// Diagnostics API/UDS/API/bds_uds_registerDidWriteCallback
///This function registers the callback for DID write operation.
///
///=======
/// Remarks:
///=======
///    + This is the mandatory API to be used if the DID parameter needs to be written.
///    + The |GVL_uds| is given for usage of defines.
///
///----------
/// FFI:
///----------
///This API can be used in trusted partitions only. See Freedom from Interference (FFI) concept for more details.
///
///==================================================================		  			===================================================================================================
///Return value    								  									Description
///==================================================================		  			===================================================================================================
///0																					No error
///1																					Invalid pointer
///
///==================================================================		   			===================================================================================================
///
///=======
///Code Example:
///=======
///============================================================================
///
///FUNCTION POU_1 : BYTE
///VAR_INPUT
///
///    can_data : POINTER TO BYTE;
///END_VAR
///
///VAR
///    data_au8 : ARRAY[0..8] OF BYTE;
///	
///    i1: BYTE;
///	
///    DidValue_u16: UINT;
///	
///    set_u8: USINT;
///END_VAR
///
///
///bds_uds_GetActiveDid(ADR(DidValue_u16));
///
///IF (DidValue_u16=16#100)
///
///  THEN bds_uds_setCallbackStatus(0);(*positive response for DID 16#100*)
///  
///END_IF
///
///IF (DidValue_u16=16#200) 
///
///  THEN  bds_uds_setCallbackStatus(1);(*negative response for DID 16#200*)
///  
///END_IF
///
///
///FOR i1 := 0 TO 8 BY 1 DO
///can_data[i1]  := data_au8[i1];
///END_FOR;
///POU_1 :=1;
///
///(*Registering callback*)
///
///PROGRAM POU_10
///VAR
///
///	flag_1 : BOOL := 1;
///	
///    flag_2 : BOOL := 1; 
///   
///    flag_3 : BOOL := 1;    
///
///END_VAR
///
///IF ( flag_1)
///
///    THEN bds_uds_registerDidReadCallback (ADR(POU_1));
///
///    flag_1 := 0;(*To make api call once in application*)
///
///END_IF
///
///IF ( flag_2)
///
///    THEN bds_uds_registerDidWriteCallback (ADR(POU_1));
///
///    flag_2 := 0;(*To make api call once in application*)
///
///END_IF
///
///IF ( flag_3)
///
///    THEN bds_uds_registerRoutineF000Callback (ADR(POU_3));
///
///    flag_3 := 0;(*To make api call once in application*)
///
///END_IF
///
///
///============================================================================
{attribute 'external_name' := 'cmp_rts_bds_uds_registerDidWriteCallback'}
FUNCTION bds_uds_registerDidWriteCallback : USINT
VAR_INPUT
	///Function pointer with argument of UINT8 data pointer
	func_pf: POINTER TO BOOL;
END_VAR

END_FUNCTION

// Diagnostics API/UDS/API/bds_uds_registerRoutineF000Callback
///This function will registers the callback for the routine control identifier F000.
///
///=======
/// Remarks:
///=======
///    + This is the mandatory API to be used for routine control identifier F000.
///	+ This is the common register API for routine control F000 for all sub functions like start(), stop(), getResults().
///    + The |GVL_uds| is given for usage of defines.
///
///----------
/// FFI:
///----------
///This API can be used in trusted partitions only. See Freedom from Interference (FFI) concept for more details.
///
///==================================================================		  			===================================================================================================
///Return value    								  									Description
///==================================================================		  			===================================================================================================
///0																					No error
///1																					Invalid pointer
///
///==================================================================		   			===================================================================================================
///
///=======
///Code Example:
///=======
///============================================================================
///
///FUNCTION POU_3 : BYTE
///VAR_INPUT
///
///    dataIn1 : BYTE;
///
///    status : BYTE;
///
///    dataOut1 : POINTER TO BYTE;
///
///    Error_Code : POINTER TO BYTE;
///
///    subservice_u8 : BYTE;
///END_VAR
///
///VAR
///    data_au8: ARRAY[0..7] OF BYTE :=[1,2,3,4,5,6,7,8];
///
///    i: BYTE;
///
///    RidValue_u16: UINT;
///
///    set: BYTE;
///END_VAR
///
///IF(subservice_u8=1)
///
///    THEN bds_uds_setCallbackStatus(0);
///
///END_IF
///
///IF(subservice_u8=2)
///
///    THEN bds_uds_setCallbackStatus(0);
///
///END_IF
///
///IF(subservice_u8=3)
///
///    THEN bds_uds_setCallbackStatus(1);
///
///END_IF
///
///(*Registering callback*)
///
///PROGRAM POU_10
///VAR
///   
///    flag_3 : BOOL := 1;    
///
///END_VAR
///
///
///IF ( flag_3)
///
///    THEN bds_uds_registerRoutineF000Callback (ADR(POU_3));
///
///    flag_3 := 0;(*To make api call once in application*)
///
///END_IF
///
///
///============================================================================
{attribute 'external_name' := 'cmp_rts_bds_uds_registerRoutineF000Callback'}
FUNCTION bds_uds_registerRoutineF000Callback : USINT
VAR_INPUT
	///Function pointer with argument of as mentioned above
	func_pf: POINTER TO BOOL;
END_VAR

END_FUNCTION

// Diagnostics API/UDS/API/bds_uds_getActiveSession
///This function gets the active session of the server/ECU.
///
///=======
/// Remarks:
///=======
///    + By default the server/ECU will be in the Default session after startup.
///    + The |GVL_uds| is given for usage of defines.
///
///----------
/// FFI:
///----------
///This API can be used in trusted partitions. For untrusted partitions use |bds_uds_getActiveSession_ffi|. See Freedom from Interference (FFI) concept for more details.
///
///==================================================================		  			===================================================================================================
///Return value    								  									Description
///==================================================================		  			===================================================================================================
///16#00																				No error
///16#01																				Invalid pointer
///16#25																				FFI API access error.
///
///==================================================================		   			===================================================================================================
///=======
///Code Example:
///=======
///============================================================================
///
///PROGRAM PLC_PRG
///  VAR
///  
///	bds_uds_session_u8:USINT;
///
///	result: USINT;
///	
///  END_VAR
///
///  (*get the active session of the ECU*)
///  
///result := bds_uds_getActiveSession(ADR(bds_uds_session_u8));
///
///============================================================================
{attribute 'external_name' := 'cmp_rts_bds_uds_getActiveSession'}
FUNCTION bds_uds_getActiveSession : USINT
VAR_INPUT
	///Reference of variable where the active session will be saved by the API. 
	///
	///The possible values are:
	///    + DEFAULT SESSION - 16#01
	///    + PROGRAMMING SESSION - 16#02
	///    + EXTENDED DIAGNOSTIC SESSION - 16#03
	///    + SAFETY SYSTEM DIAGNOSTIC SESSION - 16#04
	///    + EOL SESSION - 16#40
	bds_uds_session_u8: POINTER TO USINT;
END_VAR

END_FUNCTION

// Diagnostics API/UDS/FFI_API/bds_uds_getActiveSession_ffi
{attribute 'external_name' := 'cmp_rts_bds_uds_getActiveSession_ffi'}
FUNCTION bds_uds_getActiveSession_ffi : USINT
VAR_INPUT
	///Reference of variable where the active session will be saved by the API. 
	///
	///The possible values are:
	///    + DEFAULT SESSION - 16#01
	///    + PROGRAMMING SESSION - 16#02
	///    + EXTENDED DIAGNOSTIC SESSION - 16#03
	///    + SAFETY SYSTEM DIAGNOSTIC SESSION - 16#04
	///    + EOL SESSION - 16#40
	bds_uds_session_u8: POINTER TO USINT;
END_VAR

END_FUNCTION

// Diagnostics API/UDS/API/bds_uds_getNodeID
///This function reads the currently configured node ID, tester ID and RX/TX identifier from UDS stack and updates the input parameter.
///
///=======
/// Remarks:
///=======
///    + This function reads the UDS parameters of BODAS instance.
///    + The |GVL_uds| is given for usage of defines.
///
///----------
/// FFI:
///----------
///This API can be used in trusted partitions. For untrusted partitions use |bds_uds_getNodeID_ffi|. See Freedom from Interference (FFI) concept for more details.
///		
///==================================================================		  			===================================================================================================
///Return value    								  									Description
///==================================================================		  			===================================================================================================
///16#00																				No error
///16#01																				Node ID read failed
///16#02																				Invalid parameter
///16#25																				FFI API access error.
///
///==================================================================		   			===================================================================================================
{attribute 'external_name' := 'cmp_rts_bds_uds_getNodeID'}
FUNCTION bds_uds_getNodeID : USINT
VAR_INPUT
	///This is a union of a structure and UDINT variable.Default value : 
	///    + nodeid_u8 = 16#01
	///    + testerid_u8 = 16#FA
	///    + rxtxidentifiers_u16 = 16#18DA
	udsConfig_u: POINTER TO bds_uds_udsconfigparameter_tu;
END_VAR

END_FUNCTION

// Diagnostics API/UDS/FFI_API/bds_uds_getNodeID_ffi
{attribute 'external_name' := 'cmp_rts_bds_uds_getNodeID_ffi'}
FUNCTION bds_uds_getNodeID_ffi : USINT
VAR_INPUT
	///This is a union of a structure and UDINT variable.Default value : 
	///    + nodeid_u8 = 16#01
	///    + testerid_u8 = 16#FA
	///    + rxtxidentifiers_u16 = 16#18DA
	udsConfig_u: POINTER TO bds_uds_udsconfigparameter_tu;
END_VAR

END_FUNCTION

// Diagnostics API/UDS/API/bds_uds_permitAccess
///This function sets the access related to the BODAS-service features.
///
///=======
/// Remarks:
///=======
///    + This function needs to be called if access to the BODAS-service to be prevented/permitted.
///    + By default all the services of the BODAS-service is allowed by the BSW.
///    + Multiple bits can be set at a time.
///    + The |GVL_uds| is given for usage of defines.
///
///-----
/// DANGER:
///-----
///
///Application should take care of Programming session bit carefully.
///
///----------
/// FFI:
///----------
///This API can be used in trusted partitions only. See Freedom from Interference (FFI) concept for more details.
///
///==================================================================		  			===================================================================================================
///Return value    								  									Description
///==================================================================		  			===================================================================================================
///0																					No error
///1																					Invalid pointer
///
///==================================================================		   			===================================================================================================
///=======
///Code Example:
///=======
///============================================================================
///
///PROGRAM PLC_PRG
///  VAR
///
///	bds_uds_access_u8:USINT:=0;	
///
///	result: USINT;
///	
///  END_VAR
///  
///result:=bds_uds_permitAccess(bds_uds_access_u8);
///
///============================================================================
{attribute 'external_name' := 'cmp_rts_bds_uds_permitAccess'}
FUNCTION bds_uds_permitAccess : USINT
VAR_INPUT
	///This value defines the coded access rights for the diagnostics services of BODAS-service.
	///	
	///The supported values are:
	///    + 16#00: Prevent all services by BODAS-service.
	///    + 16#01: Permit soft reset by BODAS-service.
	///    + 16#02: Permit hard reset by BODAS-service.
	///    + 16#04: Permit keyOffOn reset by BODAS-service.
	///    + 16#10: Permit to programming session by BODAS-service.
	///    + 16#FF: Permit all services by BODAS-service. (Default)
	bds_uds_access_u8: USINT;
END_VAR

END_FUNCTION

// Diagnostics API/UDS/API/bds_uds_registerRoutineCtrlCallback
///This function will registers the callback for the any routine control configured in easyConfig.
///
///=======
/// Remarks:
///=======
///    + This API is not used for routine control identifier F000. see |bds_uds_registerRoutineF000Callback|
///	+ This is the common register API for all routine control for all sub functions like start(), stop(), getResults().
///    + The |GVL_uds| is given for usage of defines.
///
///----------
/// FFI:
///----------
///This API can be used in trusted partitions only. See Freedom from Interference (FFI) concept for more details.
///
///==================================================================		  			===================================================================================================
///Return value    								  									Description
///==================================================================		  			===================================================================================================
///0																					No error
///1																					Invalid pointer
///
///==================================================================		   			===================================================================================================
///
///=======
///Code Example:
///=======
///============================================================================
///
///FUNCTION POU_3 : BYTE
///VAR_INPUT
///
///    dataIn1 : POINTER TO BYTE;
///
///    status : BYTE;
///
///    dataOut1 : POINTER TO BYTE;
///
///    Error_Code : POINTER TO BYTE;
///
///	(*subservice not available for this function*)
///
///END_VAR
///
///VAR
///    data_au8: ARRAY[0..7] OF BYTE :=[1,2,3,4,5,6,7,8];
///
///    i: BYTE;
///
///    RidValue_u16: UINT;
///
///    set: BYTE;
///END_VAR
///
///IF(subservice_u8=1) THEN
///
///     bds_uds_setCallbackStatus(0);
///
///END_IF
///
///IF(subservice_u8=2) THEN
///
///     bds_uds_setCallbackStatus(0);
///
///END_IF
///
///IF(subservice_u8=3) THEN
///
///     bds_uds_setCallbackStatus(1);
///
///END_IF
///
///(*Registering callback*)
///
///PROGRAM POU_10
///VAR
///   
///    flag_3 : BOOL := 1;    
///
///END_VAR
///
///
///IF ( flag_3)
///
///    THEN bds_uds_registerRoutineCtrlCallback (ADR(POU_3));
///
///    flag_3 := 0;(*To make api call once in application*)
///
///END_IF
///
///
///============================================================================
{attribute 'external_name' := 'cmp_rts_bds_uds_registerRoutineCtrlCallback'}
FUNCTION bds_uds_registerRoutineCtrlCallback : USINT
VAR_INPUT
	///Function pointer with argument as mentioned above
	func_pf: POINTER TO BOOL;
END_VAR

END_FUNCTION

// I/O API/OUT_LEGACY/bds_out_po_disableTstPls
///Disables test pulses for a dedicated proportional output to avoid having test pulses for error detection on that output.
///
///=======
/// Remarks:
///=======
///
///   + Test pulses are enabled by default.
///   + For some application the test pulses may disturb the required functionality of an output. For example if you want to use it for power supply.
///   + The test pulses can be deactivated for High Power Outputs only.
///   + This function should be called only once in the application.
///
///----------
/// FFI:
///----------
///This API can be used in trusted partitions . For untrusted partitions use |bds_out_po_disableTstPls_ffi|. See Freedom from Interference (FFI) concept for more details.
///
///------
/// Attention:
///------
///
///If test pulses are disabled for an output, fault detection and healing is limited.
///
///==================================================================		  			===================================================================================================
///Return value    								  									Description
///==================================================================		  			===================================================================================================
///0																					No error.
///1																					Signal is out of range.
///2																					State Command out of range.
///3																					Output is configured as safout, Test pulse can't be disabled
///
///==================================================================		   			===================================================================================================
///
///=======
///Code Example:
///=======
///============================================================================
///
///PROGRAM PLC_PRG
///
///VAR
///
///	Init_flag_u8:USINT:=0;
///
///END_VAR
///  
///IF(Init_flag_u8=0) THEN (*To make api call once in application*)
///				
///	(* disable test pulses for output K07 *)
///	
///	bds_out_po_disableTstPls(bds_out_po_signal_te.K07, STD_ON);
///  
///	Init_flag_u8:=1;
///  
///END_IF
///
///============================================================================
{attribute 'external_name' := 'cmp_rts_bds_out_po_disableTstPls'}
FUNCTION bds_out_po_disableTstPls : USINT
VAR_INPUT
	///The connector assigned signal name of the output.
	signal_e: UINT;
	///The states are
	///   + STD_OFF - Enables the test pulses (default)
	///   + STD_ON   - Disables the test pulses
	state_u8: USINT;
END_VAR

END_FUNCTION

// I/O API/OUT/FFI_API/bds_out_po_disableTstPls_ffi
{attribute 'external_name' := 'cmp_rts_bds_out_po_disableTstPls_ffi'}
FUNCTION bds_out_po_disableTstPls_ffi : USINT
VAR_INPUT
	///The connector assigned signal name of the output.
	signal_e: UINT;
	///The states are
	///   + STD_OFF - Enables the test pulses (default)
	///   + STD_ON   - Disables the test pulses
	state_u8: USINT;
END_VAR

END_FUNCTION

// I/O API/OUT_LEGACY/bds_out_po_getCurrent
///Get the current of the proportional output.
///
///=======
/// Remarks:
///=======
///   + The threshold for the over current detection is 6000mA and therefore also the measurement range is defined from 0..6000mA.
///
///----------
/// FFI:
///----------
///This API can be used in trusted partitions . For untrusted partitions use |bds_out_po_getCurrent_ffi|. See Freedom from Interference (FFI) concept for more details.
///
///==================================================================		  			===================================================================================================
///Return value    								  									Description
///==================================================================		  			===================================================================================================
///0																					No error.
///1																					A parameter is invalid.
///2																					Function call was erroneous.
///
///==================================================================		   			===================================================================================================
///
///=======
///Code Example:
///=======
///============================================================================
///
///PROGRAM appl_10ms_task
///VAR
///bds_outClcU_signal_e : bds_outClcU_signal_te;
/// bds_outClcU_retSetVoltage_s : bds_outClcU_setVoltage_ts;
/// u_mV_u16 : UINT := 8000;
///END_VAR
///
///bds_outClcU_signal_e := bds_outClcU_K62_E;
///
///bds_outClcU_retSetVoltage_s := bds_outClcU_setVoltage(bds_outClcU_signal_e, u_mV_u16);
///
///IF bds_outCmn_ok_E = bds_outClcU_retSetVoltage_s.statusApi_e THEN
/// (* Call successful, signal is valid )
/// ( Set point value is set on requested output )
///  ELSE
///  ( error handling *)
///  END_IF
///
///END_PROGRAM
///============================================================================
{attribute 'external_name' := 'cmp_rts_bds_out_po_getCurrent'}
FUNCTION bds_out_po_getCurrent : USINT
VAR_INPUT
	///The connector assigned signal name of the output.
	signal_e: UINT;
	///Storage address of the value.
	///
	///   + Range:0 to 60000 [mA]
	value_pu16: POINTER TO UINT;
END_VAR

END_FUNCTION

// I/O API/OUT/FFI_API/bds_out_po_getCurrent_ffi
{attribute 'external_name' := 'cmp_rts_bds_out_po_getCurrent_ffi'}
FUNCTION bds_out_po_getCurrent_ffi : USINT
VAR_INPUT
	///The connector assigned signal name of the output.
	signal_e: UINT;
	///Storage address of the value.
	///
	///   + Range:0 to 60000 [mA]
	value_pu16: POINTER TO UINT;
END_VAR

END_FUNCTION

// I/O API/OUT/API/bds_outClcU_setVoltage
///The BODAS API-Function sets the analog voltage set point of the output signal.
///
///=======
/// Remarks:
///=======
///    +For AOV analog voltage output the set voltage range is from 0 to 10000mV  (available signal refer to table "AOV Analog Voltage Output" in RC27-18/40 - Outputs).
///    
///    +For PVG proportional voltage output the accepted set voltage range is from 0 to 27000mV (75% of max Ubat) (available signal refer to table "PVG Proportional Voltage Output" in RC27-18/40 - Outputs).
///   
///    +·If the set point has been set to 0 value then the output can also be used as analog voltage input, refer to bds_outClcU_get.
///
///----------
/// FFI:
///----------
///This API can be used in trusted partitions. For untrusted partitions use bds_outClcU_setVoltage_ffi. See Freedom from Interference (FFI) concept for more details.
///
///------
/// Info:
///------
///
/// +For the output type PVG: 
///   
///   +An external load is mandatory, refer to Technical Data Sheet (RE-sheet RE95207).
///   
///   +If the requested voltage set point is higher than 75% of the max possible battery voltage (36V) the return value of the status API function call is: bds_outCmn_outOfRng_E.
///   
///   +·The possible voltage range that can be controlled is 25% to 75% of the actual battery voltage, because of hardware limitations. The internal set point of the regulation will be dynamically limited to this min or max value without setting any error or status information.
///
///   +Example 1: 
///   +Actual battery voltage = 24V and output voltage is set to 4V => results in output voltage = 6V (25% of actual battery voltage).
///
///   +Example 2: 
///   +Actual battery voltage = 12V and output voltage is set to 4V => results in output voltage = 4V (33% of actual battery voltage).
///   
///   +The set point request of 0V is also valid and will switch off the output. 
///   
///   
///   +Macro define "bds_outClcU_strtNumSigAov_D" in easyConfig generated file "bds_outClcU_ec.h" defines the start of the Analog voltage output (AOV) signals in the enumeration type definition "bds_outClcU_signal_te".
///
///
///==================================================================		  			===================================================================================================
///Return value    								  									Description
///==================================================================		  			===================================================================================================
///bds_outClcU_setVoltage_ts															 The return structure containing the state information (statusApi_e)
///
///==================================================================		   			===================================================================================================
///
///=======
///Code Example:
///=======
///============================================================================
///
///PROGRAM appl_10ms_task
///
///VAR
///
///bds_outClcU_signal_e : bds_outClcU_signal_te;
///
///bds_outClcU_retSetVoltage_s : bds_outClcU_setVoltage_ts;
///
///u_mV_u16 : UINT := 8000;
///
///END_VAR
///
///bds_outClcU_signal_e := bds_outClcU_signal_te.bds_outClcU_K62_E;
///
///bds_outClcU_retSetVoltage_s := bds_outClcU_setVoltage(bds_outClcU_signal_e, u_mV_u16);
///
///IF bds_outCmn_ok_E = bds_outClcU_retSetVoltage_s.statusApi_e THEN
///
///(* Call successful, signal is valid *)
///(* Set point value is set on requested output *)
///
///ELSE
///
///(* error handling *)
///
///END_IF
///
///END_PROGRAM
///
///============================================================================
{attribute 'external_name' := 'cmp_rts_bds_outClcU_setVoltage'}
FUNCTION bds_outClcU_setVoltage : bds_outClcU_setVoltage_ts
VAR_INPUT
	///signal name of the output (connector pin)
	signal_e: USINT;
	///New set point for PWM [0.1%] respective AOV [mV].Range:
	///   + PWM: 0 and 250 to 750
	///   + AOV: 0 to 10000
	u_mV_u16: UINT;
END_VAR

END_FUNCTION

// I/O API/OUT/API/bds_outClcU_get
///The BODAS API-Function gets the measured voltage in [mV] of the analog voltage output pin.
///
///=======
/// Remarks:
///=======
///  +The voltage range depends on the type.
/// 
///     +AOV: 0 to 12000mV
/// 
///     +PVG: 0 to 33000mV.
/// 
///  +The read-back path of the analoge voltage can also be used as analog input, if the set point is set to zero, refer also bds_outClcU_setVolatge and bds_outClcU_setPercUBat.
///  +Diagnostics capabilities similar to standard inputs is not available. 
/// 
///  +The status data holds all relevant information of the analog voltage output, see example below.
/// 
///  +Part of the status bit field is also the fault error status of every DFC (e.g. stErrSCB_b1), see topic Digital outputs and Diagnostic Fault Check. 

///
///----------
/// FFI:
///----------
///This API can be used in both trusted and untrusted partitions. See Freedom from Interference (FFI) concept for more details.
///
///------
/// Info:
///------
///
///   +For the predefined pin type analog voltage output (AOV) there is an option in easyConfig tool to reconfigure it as analog voltage input or digital input
///
///
///==================================================================		  			===================================================================================================
///Return value    								  									    Description
///==================================================================		  			===================================================================================================
///bds_outClcU_get_ts															        The return structure containing the measured voltage in [mV] and the state information (statusApi_e)
///
///==================================================================		   			===================================================================================================
///
///=======
///Code Example:
///=======
///============================================================================
///
/// PROGRAM appl_10ms_task 
///
/// VAR
/// 
/// bds_outClcU_signal_e : bds_outClcU_signal_te; 
/// 
/// bds_outClcU_retGet_s : bds_outClcU_get_ts; 
///
/// retVal_uAct_mV_u16, retVal_uSet_mV_u16 : UINT;
/// 
/// END_VAR
///
/// bds_outClcU_signal_e := bds_outClcU_signal_te.bds_outClcU_K62_E; 
///
///
/// (* call BDS-Function - Set voltage output *)
///
/// bds_outClcU_setVoltage(bds_outClcU_signal_e, 8000); 
///
/// (* call BDS-Function - Get status and diagnostic information *)
///
/// bds_outClcU_retGet_s := bds_outClcU_get(bds_outClcU_signal_e); 
///
///
/// IF bds_outCmn_ok_E = bds_outClcU_retGet_s.statusApi_e THEN
///
/// (* Call successful, signal is valid *)
///
/// 	(* check if there is a short cut to battery or to ground? *)
///
///		IF (TRUE = bds_outClcU_retGet_s.statusDiag_b.stErrSCB_b1) OR (TRUE = bds_outClcU_retGet_s.statusDiag_b.stErrSCG_b1) THEN
///
/// 	(* SCB or SCG - Set values to zero *)
///
///  	retVal_uAct_mV_u16 := 0; 
///
/// 	retVal_uSet_mV_u16 := 0; 
///
/// 	ELSE (* get actual measured voltage on requested output *)
///
///		retVal_uAct_mV_u16 := bds_outClcU_retGet_s.uAct_mV_u16; 
///
///     (* get requested set point voltage on requested output *)
///
///     retVal_uSet_mV_u16 := bds_outClcU_retGet_s.uSet_mV_u16; 
///
/// 	END_IF
///
/// ELSE
///
/// (* error handling *)
///
/// END_IF
///
/// END_PROGRAM
///
///============================================================================
{attribute 'external_name' := 'cmp_rts_bds_outClcU_get'}
FUNCTION bds_outClcU_get : bds_outClcU_get_ts
VAR_INPUT
	///signal name of the output (connector pin)
	signal_e: USINT;
END_VAR

END_FUNCTION

// I/O API/OUT/API/bds_outClcU_setPercUBat
/// The BODAS API-Function sets the analog voltage output in percentage value of the the battery voltage.
///
///=======
/// Remarks:
///=======
///    +Set the voltage range FROM 0 AND 250…750 [0.1%] OF the battery voltage OF the PVG analog voltage output (available signal refer TO table "PVG Proportional Voltage Output" in RC27-18/40 - Outputs).

///    +If the set point has been set to 0 value then the output can also be used as analog voltage input, refer to bds_outClcU_get.

///
///----------
/// FFI:
///----------
/// This API can be used in trusted partitions. For untrusted partitions use bds_outClcU_setPercUBat_ffi. See Freedom from Interference (FFI) concept for more details.
///
///------
/// Info:
///------
///
/// +For the output type PVG an external load is mandatory, refer to Technical Data Sheet (RE-sheet RE95207).
/// +Macro define "bds_outClcU_strtNumSigAov_D" in easyConfig generated file "bds_outClcU_ec.h" defines the start of the Analog voltage output (AOV) signals in the enumeration type definition "bds_outClcU_signal_te"
///
///
///==================================================================		  			===================================================================================================
///Return value    								  									    Description
///==================================================================		  			===================================================================================================
///bds_outClcU_setPercUBat_ts														     The return structure containing the state information (statusApi_e)
///
///==================================================================		   			===================================================================================================
///
///=======
///Code Example:
///=======
///============================================================================
///
/// PROGRAM appl_10ms_task 
///
/// VAR bds_outClcU_signal_e : bds_outClcU_signal_te;
///
/// bds_outClcU_retSetPercUBat_s : bds_outClcU_setPercUBat_ts;
///
/// ratUBat_perml_u16 : UINT;
///
/// END_VAR
///
/// bds_outClcU_signal_e := bds_outClcU_signal_te.bds_outClcU_K25_E;
///
/// ratUBat_perml_u16 := 750;
///
///bds_outClcU_retSetPercUBat_s := bds_outClcU_setPercUBat(bds_outClcU_signal_e, ratUBat_perml_u16);
///
///IF bds_outCmn_ok_E = bds_outClcU_retSetPercUBat_s.statusApi_e THEN 
///
/// (* Call successful, signal is valid *)
///
/// (* Set point value is set on requested output *)
///
/// ELSE
/// 
/// (* error handling *)
///
/// END_IF
///
/// END_PROGRAM
///
///============================================================================
{attribute 'external_name' := 'cmp_rts_bds_outClcU_setPercUBat'}
FUNCTION bds_outClcU_setPercUBat : bds_outClcU_setPercUBat_ts
VAR_INPUT
	///signal name of the output (connector pin)
	signal_e: USINT;
	///voltage set point in 0, 250...750 [0.1%] of battery voltage
 
	ratUBat_perml_u16: UINT;
END_VAR

END_FUNCTION

// Diagnostics API/UDS/API/bds_uds_setUUID
///This function is to set the Universal Unique Identifier for ODX file data identification.
///
///=======
/// Remarks:
///=======
///
///    + UDS dataidentifier 16#F19E supports the UUID-ODX data identification value set from |bds_uds_setUUID|.
///    + The |GVL_uds| is given for usage of defines.
///    + This API should be called once in Application
///
///----------
/// FFI:
///----------
///This API can be used in trusted partitions only. See Freedom from Interference (FFI) concept for more details.
///
///----------
/// WARNING:
///----------
///
///This function should be called only once in the application.
///
///==================================================================		  			===================================================================================================
///Return value    								  									Description
///==================================================================		  			===================================================================================================
///16#00																				No error
///16#01																				Invalid pointer
///
///==================================================================		   			===================================================================================================
///=======
///Code Example:
///=======
///============================================================================
///
///PROGRAM PLC_PRG
///  VAR
///
///	bds_uds_uuid_pu8: ARRAY[0 .. 17] OF USINT;
///
///	bds_uds_uuidLen_u8 : USINT := 18;
///
///	result: USINT;
///
///	FLAG: BOOL;
///	
///  END_VAR
///  
///IF FLAG:=FALSE THEN
///
///	bds_uds_uuid_pu8[0]:= 16#FF; 
///
///	bds_uds_uuid_pu8[1]:= 16#AA; 
///
///	result := bds_uds_setUUID(ADR(bds_uds_uuid_pu8),bds_uds_uuidLen_u8);
///
///	FLAG:= TRUE;
///
///END_IF
///
///============================================================================
{attribute 'external_name' := 'cmp_rts_bds_uds_setUUID'}
FUNCTION bds_uds_setUUID : USINT
VAR_INPUT
	///Array index for the 18 byte UUID value for ODX identification
	bds_uds_uuid_pu8: POINTER TO USINT;
	///Length in bytes for the UUID value, maximum is 18.
	bds_uds_uuidLen_u8: USINT;
END_VAR

END_FUNCTION

// I/O API/SAFOUT/API/bds_safout_cfgDiag
///Configures the allowed current deviation limit for current deviation monitoring between high side and low side outputs of a safout channel. 
///
///=======
/// Remarks:
///=======
///   + The allowed default current deviation limit is 100 mA. Current deviation monitoring between high side and low side outputs is supported only for PHMDL, PLMDH, PLDHS and PHDLS mode.
///   + Some of the errors are detected using current deviation monitoring, setting of allowed current deviation limit shall be chosen wisely for the application. 
///   + Total allowed current deviation limit = (Current deviation in mA + (percentage of sum of current through multiple side outputs in previous100 ms) in mA).
///
///----------
/// FFI:
///----------
///This API can be used in trusted partitions only. See Freedom from Interference (FFI) concept for more details.
///
///------
/// CAUTION:
///------
///
///Be careful while configuring current deviation.
///
///==================================================================		  			===================================================================================================
///Return value    								  									Description
///==================================================================		  			===================================================================================================
///0																					No error
///1																					A parameter is invalid
///2																					Wrong mode or channel
///3																					Feature not supported for safout mode
///
///==================================================================		   			===================================================================================================
///
///=======
///Code Example:
///=======
///============================================================================
///
///VAR_GLOBAL CONSTANT
///
///   (* safout channel name *)
///
///   PHDLS_CHNL1: UINT := (PHDLS OR CHNL1);
///
///   DHDLM_CHNL2: UINT := (DHDLM OR CHNL2);
///
///   PHMDL_CHNL3: UINT := (PHMDL OR CHNL3);
///   
///   PLDHS_CHNL4: UINT := (PLDHS OR CHNL4);
///
///   DLDHM_CHNL5: UINT := (DLDHM OR CHNL5);
///
///   PLMDH_CHNL6: UINT := (PLMDH OR CHNL6);
///
///END_VAR
///
///PROGRAM PLC_PRG
///
///VAR
///
///END_VAR
///
///
///(* configure for POC *)
///
///bds_out_po_cfg(bds_out_po_signal_te.K73, STD_ACTIVE);
///
///bds_out_po_cfg(bds_out_po_signal_te.K07, STD_ACTIVE);
///
///bds_out_po_cfg(bds_out_po_signal_te.K29, STD_ACTIVE);
///
///bds_out_po_cfg(bds_out_po_signal_te.K09, STD_ACTIVE);
///
///
///
///(* configure channels for SAFOUT *)
///
///bds_safout_cfg(PHDLS_CHNL1, bds_out_po_signal_te.K73, bds_out_po_signal_te.K51, bds_out_do_signal_te.K14, 0, 0);
///
///bds_safout_cfg(DHDLM_CHNL2, bds_out_po_signal_te.K08, bds_out_do_signal_te.K16, bds_out_do_signal_te.K15, bds_out_do_signal_te.K13, 0);
///
///bds_safout_cfg(PHMDL_CHNL3, bds_out_do_signal_te.K12, bds_out_po_signal_te.K07, bds_out_po_signal_te.K29, bds_out_po_signal_te.K09, 0);
///
///bds_safout_cfg(PLDHS_CHNL4, bds_out_po_signal_te.A19, bds_out_po_signal_te.A32, bds_out_do_signal_te.A47, 0, 0);
///
///bds_safout_cfg(DLDHM_CHNL5, bds_out_po_signal_te.A03, bds_out_do_signal_te.A33, bds_out_do_signal_te.A46, bds_out_do_signal_te.A48, 0);
///
///bds_safout_cfg(PLMDH_CHNL6, bds_out_do_signal_te.A31, bds_out_po_signal_te.A05, bds_out_po_signal_te.A20, 0, 0);
///
///bds_safout_cfgDiag(PHDLS_CHNL1, 150,0);
///
///bds_safout_cfgDiag(PHMDL_CHNL3, 200, 10);
///
///bds_safout_cfgDiag(PLDHS_CHNL4, 200,15);
///
///bds_safout_cfgDiag(PLMDH_CHNL6, 200, 10);
///
///============================================================================
{attribute 'external_name' := 'cmp_rts_bds_safout_cfgDiag'}
FUNCTION bds_safout_cfgDiag : USINT
VAR_INPUT
	///The connector assigned signal name of the output.
	///
	///The channel name is composed of mode and channel number
	///
	///channel name = mode OR channel number
	///
	///and shall be defined from the application (see also example below):
	///
	///PHDLS_CHNL1: UINT := (PHDLS OR CHNL1)
	chnl_u16: UINT;
	///Fixed allowed current deviation [mA] 
	///   + Range: 100..1000 
	deviation_u16: UINT;
	///Percentage of allowed current deviation [%]
	///   + Range:0..100
	devPercentage_u8: USINT;
END_VAR

END_FUNCTION

// I/O API/SAFOUT/API/bds_safout_enableTest
///Enables test for Safout channel.
///
///When safout channel is inactive i.e all highsides and lowside are OFF, every 2 seconds a test is performed by switching ON common side for 120 ms.  During test, open load error diagnostic is performed on multiple outputs of the safout channel can be detected.
///
///=======
/// Remarks:
///=======
///   + A channel shall be configured with ECU specific modes, see Safety outputs.
///   + By default, test is disabled 
///   + This test is not performed when there a SCB on HS output / SCG on LS outputs.
///   + Test status can be using |bds_safout_getStatus| API. Test complete flag is reset once status is read by |bds_safout_getStatus|.
///   + This only supported for PHMDL mode. In other safout modes open load is detected without this test.
///
///----------
/// FFI:
///----------
///This API can be used in trusted partitions only. See Freedom from Interference (FFI) concept for more details.
///
///==================================================================		  			===================================================================================================
///Return value    								  									Description
///==================================================================		  			===================================================================================================
///0																					No error.
///1																					A parameter is invalid.
///2																					Not supported for this mode
///
///==================================================================		   			===================================================================================================
///
///=======
///Code Example:
///=======
///============================================================================
///
///VAR_GLOBAL CONSTANT
///
///   (* safout channel name *)
///
///   PHDLS_CHNL1: UINT := (PHDLS OR CHNL1);
///
///   DHDLM_CHNL2: UINT := (DHDLM OR CHNL2);
///
///   PHMDL_CHNL3: UINT := (PHMDL OR CHNL3);
///
///END_VAR
///
///PROGRAM PLC_PRG
///
///VAR
///
///END_VAR
///
///(* configure for POC *)
///
///bds_out_po_cfg(bds_out_po_signal_te.K73, STD_ACTIVE);
///
///bds_out_po_cfg(bds_out_po_signal_te.K07, STD_ACTIVE);
///
///bds_out_po_cfg(bds_out_po_signal_te.K29, STD_ACTIVE);
///
///bds_out_po_cfg(bds_out_po_signal_te.K09, STD_ACTIVE);
///
///
///(* configure channels for SAFOUT *)
///
///bds_safout_cfg(PHDLS_CHNL1, bds_out_po_signal_te.K73, bds_out_po_signal_te.K51, bds_out_do_signal_te.K14, 0, 0);
///
///bds_safout_cfg(DHDLM_CHNL2, bds_out_po_signal_te.K08, bds_out_do_signal_te.K16, bds_out_do_signal_te.K15, bds_out_do_signal_te.K13, 0);
///
///bds_safout_cfg(PHMDL_CHNL3, bds_out_do_signal_te.K12, bds_out_po_signal_te.K07, bds_out_po_signal_te.K29, bds_out_po_signal_te.K09, 0);
///
///bds_safout_enableTest(PHMDL_CHNL3,STD_ON);
///
///============================================================================
{attribute 'external_name' := 'cmp_rts_bds_safout_enableTest'}
FUNCTION bds_safout_enableTest : USINT
VAR_INPUT
	///The connector assigned signal name of the output.
	///
	///The channel name is composed of mode and channel number
	///
	///channel name = mode OR channel number
	///
	///and shall be defined from the application (see also example below):
	///
	///PHDLS_CHNL1: UINT := (PHDLS OR CHNL1)
	chnl_u16: UINT;
	///The states are
	///   + STD_OFF - Disable the test (default)
	///   + STD_ON   - Enable the test
	state_u8: USINT;
END_VAR

END_FUNCTION

// I/O API/IN legacy/API/bds_in_ri_cfg
///Configures the diagnosis threshold resistances for an input. 
///
///=======
/// Remarks:
///=======
///   + The information about definitions and structures can be found in BODAS API library and  bds_rts_ec.xml.
///   + The diagnosis of the input is only possible after the configuration of the thresholds.
///   + With a defined measurement range of 20 to 400k ohm the diagnosis range is defined from 30 to 399.99k ohm.
///   + For more information see |bds_in_ri_getStatus|.
///   + This function should be called only once in the application.
///
///
///----------
/// FFI:
///----------
///This API can be used in trusted partitions only. See Freedom from Interference (FFI) concept for more details.
///
///==================================================================		  			===================================================================================================
///Return value    								  									Description
///==================================================================		  			===================================================================================================
///0																					No error
///1																					Invalid parameter
///2																					Function call was erroneous
///
///==================================================================		   			===================================================================================================
///
///
///=======
///Code Example:
///=======
///============================================================================
///
///PROGRAM PLC_PRG
///
///  VAR
///  
///	Init_flag_u8:USINT:=0;
/// 
///  END_VAR
///  
///IF(Init_flag_u8=0) THEN (*To make api call once in application*)
///
///	(* configure diagnosis thresholds of input K60 *)
///	
///	bds_in_ri_cfg(bds_in_ri_signal_te.K60, 2000, 200);
///	
///	Init_flag_u8:=1;
///  
///END_IF
///
///============================================================================
{attribute 'external_name' := 'cmp_rts_bds_in_ri_cfg'}
FUNCTION bds_in_ri_cfg : USINT
VAR_INPUT
	///The signal name that is assigned to the respective pin configured as resistance input
	signal_e: UINT;
	///Upper diagnosis threshold [ohm].
	///
	///Range: 
	///30 to 399990
	///
	///Note:
	///upperThreshold_u32 > lowerThreshold_u32.  
	upperThreshold_u32: UDINT;
	///Lower diagnosis threshold [ohm].
	///
	///Range: 
	///30 to 399990
	///
	///Note:
	///lowerThreshold_u32 < upperThreshold_u32 
	lowerThreshold_u32: UDINT;
END_VAR

END_FUNCTION

// I/O API/IN legacy/API/bds_in_ri_getStatus
///Provides the status of an input.
///
///=======
/// Remarks:
///=======
///   + For information about the signal acquisition see Analog voltage aquisition.
///   + The status data provides all relevant information of the resistance input.  See the example below.
///	   + A member variable  of  the status data structure  provides the fault status of corresponding  DFC (e.g., stDFC_SCB_u16), see topic Diagnostic Fault Check. 
///	   + With the macros (e.g., bds_dsm_DFC_ldf) defined in bds_dsm_api.h  respective bit fields of the fault status can be read.
///
///----------
/// FFI:
///----------
///This API can be used in trusted partitions only. See Freedom from Interference (FFI) concept for more details.
///
///==================================================================		  			===================================================================================================
///Return value    								  									Description
///==================================================================		  			===================================================================================================
///0																					No error
///1																					Invalid parameter
///
///==================================================================		   			===================================================================================================
///
///=======
///Code Example:
///=======
///============================================================================
///
///PROGRAM appl_10ms_task
///  VAR
///  
///    stK60_s: bds_in_ri_ts;
///	
///    ldf_u8: USINT := 16#00;
///	
///  END_VAR
///
///
///(* get the status of input K60 *)
///
///bds_in_ri_getStatus(bds_in_ri_signal_te.K60, ADR(stK60_s));
///
///  (* get last debounced fault *)
///  
///  ldf_u8 = bds_dsm_DFC_ldf(stK60_s.stDFC_SCB_u16);
///END
///
///============================================================================
{attribute 'external_name' := 'cmp_rts_bds_in_ri_getStatus'}
FUNCTION bds_in_ri_getStatus : USINT
VAR_INPUT
	///The signal name that is assigned to the respective pin configured as resistance input
	signal_e: UINT;
	///Storage address of the data
	data_ps: POINTER TO bds_in_ri_ts;
END_VAR

END_FUNCTION

// I/O API/IN legacy/API/bds_in_ri_cfgTemp
///Configures the resistance inputs for temperature measurement. 
///
///=======
/// Remarks:
///=======
///   + The supported BSW sensors are:
///	   + TSF (sensor type is PTC) 
///	   + TSA (sensor type is PTC)
///	   + TFW (sensor type is NTC)
///   + For additional sensors the corresponding look up tables shall be defined, for more information see Define a look up table for temperature sensors.
///
///
///----------
/// FFI:
///----------
///This API can be used in trusted partitions only. See Freedom from Interference (FFI) concept for more details.
///
///
///==================================================================		  			===================================================================================================
///Return value    								  									Description
///==================================================================		  			===================================================================================================
///0																					No error
///1																					Invalid parameter
///
///==================================================================		   			===================================================================================================
///
///
///=======
///Code Example:
///=======
///============================================================================
///
///PROGRAM PLC_PRG
///
///  VAR
///  
///    lookup_TSF_cau16: ARRAY[1..256] OF UINT := [256(0)];
///	
///    lookup_TSA_cau16: ARRAY[1..256] OF UINT := [256(0)];
///	
///    lookup_TFW_cau16: ARRAY[1..256] OF UINT := [256(0)];
///	
///	Init_flag_u8:USINT:=0;
///	
///  END_VAR
///  
///IF(Init_flag_u8=0) THEN (*To make api call once in application*)
///
///	(* configure temperature sensor of input K60 *)
///	
///	bds_in_ri_cfgTemp(bds_in_ri_signal_te.K60, lookup_TSF_cau16, PTC);
///	
///	bds_in_ri_cfgTemp(bds_in_ri_signal_te.K58, lookup_TFW_cau16, NTC);
///	
///	Init_flag_u8:=1;
///  
///END_IF
///
///============================================================================
{attribute 'external_name' := 'cmp_rts_bds_in_ri_cfgTemp'}
FUNCTION bds_in_ri_cfgTemp : USINT
VAR_INPUT
	///The signal name that is assigned to the respective pin configured as resistance input
	signal_e: UINT;
	///Predefined look up tables for the BODAS-BSW are:
	///   + lookup_TSF_cau16 
	///   + lookup_TSA_cau16
	///   + lookup_TFW_cau16
	lookup_pcau16: POINTER TO UINT;
	///Selected sensor type are:
	///   + NTC 
	///   + PTC 
	type_u8: USINT;
END_VAR

END_FUNCTION

// I/O API/IN legacy/API/bds_in_sent_getSDDatabox
///It provides the oldest slow serial data from a particular databox of a particular SENT channel.
///
///=======
/// Remarks:
///=======
///   + The receive databoxes must be registered with |bds_in_sent_registerSDDataboxes| and then the specific receive databox has to be initialized by |bds_in_sent_initSDDatabox|.
///   + The return value  should be checked first before accessing the data/message.
///
/// 
///----------
/// FFI:
///----------
///This API can be used in trusted partitions only. See Freedom from Interference (FFI) concept for more details.
/// 
///==================================================================		  			===================================================================================================
///Return value    								  									Description
///==================================================================		  			===================================================================================================
///0																					No error
///1																					Invalid parameter
///2																					Databox is not initialized
///3																					Receive buffer is empty
///4																					Receive buffer overflow
///
///==================================================================		   			===================================================================================================
///
///=======
///Code Example:
///=======
///============================================================================
///
///VAR_GLOBAL CONSTANT
///
///   SENT_NUM_DATABOXES_D: USINT := 5;
///
///   SENT_DATABOX_BUFLEN_D: UDINT := 10;
///
///END_VAR
///
/// 
///
///PROGRAM PLC_PRG
///
///   VAR
///
///     sent_dataBox_as: ARRAY[1..SENT_NUM_DATABOXES_D] OF bds_in_sent_SDDataBox_ts;
///
///     sent_slowData1_as: ARRAY[1..SENT_DATABOX_BUFLEN_D] OF bds_in_sent_slowData_ts;
///
///     databoxdata_au16: ARRAY[1..SENT_NUMOFDATABOX_D] OF UINT;
///	 
///	Init_flag_u8:USINT:=0;	 
///
///   END_VAR
///  
///IF(Init_flag_u8=0) THEN (*To make api call once in application*)
///
///   (* register slow databox *)
///
///   bds_in_sent_registerSDDataboxes(bds_in_sent_signal_te.K52, ADR(sent_dataBox_as), SENT_NUM_DATABOXES_D);
///
/// 
///
///   (* initialize the databox *)
///
///   bds_in_sent_initSDDatabox(bds_in_sent_signal_te.K52, 1, 2, ADR(sent_slowData1_as), 5);
///	
///	Init_flag_u8:=1;
///  
///END_IF
///
/// 
///
///PROGRAM appl_10ms_task
///
///  uint8 statusSDDatabox_u8;
///
///  statusSDDatabox_u8 := bds_in_sent_getSDDatabox(bds_in_sent_signal_te.K52,1, &databoxdata_au16[0]);
///
/// 
///
///  IF (0 = statusSDDatabox_u8) THEN
///
///    (* valid data box of SLOW data *)
///
///  END_IF
///
///END
///
///
///============================================================================
{attribute 'external_name' := 'cmp_rts_bds_in_sent_getSDDatabox'}
FUNCTION bds_in_sent_getSDDatabox : USINT
VAR_INPUT
	///The signal name that is assigned to the respective pin configured as SENT input
	signal_e: UINT;
	///Number of data box
	numDatabox_u8: USINT;
	///Pointer to data array
	data_pu16: POINTER TO UINT;
END_VAR

END_FUNCTION

// I/O API/IN legacy/API/bds_in_sent_registerSDDataboxes
///The function registers a slow Databox for a particular message of particular SENT channel. Application has to reserve the memory for databox and databox is managed by the BODAS-BSW.
///
///=======
/// Remarks:
///=======
///
///   + Receive databoxes which has to be registered with function described. Each receive databox has to be initialized with function |bds_in_sent_initSDDatabox|.
///   + The use of receive databoxes is optional.
///   + By default no databoxes are registered. 
///   + For each SENT channel seperate receive databoxes must be registered. 
///   + Please register receive databoxes only as much as needed. Each receive databox increases the system load (if a SENT message is received). 
/// 
///
///----------
/// FFI:
///----------
///This API can be used in trusted partitions only. See Freedom from Interference (FFI) concept for more details.
///
///==================================================================		  			===================================================================================================
///Return value    								  									Description
///==================================================================		  			===================================================================================================
///0																					No error
///1																					Invalid parameter
///2																					new buffer overlaps a present buffer
///
///==================================================================		   			===================================================================================================
///
///=======
///Code Example:
///=======
///============================================================================
///
///VAR_GLOBAL_CONSTANT
///
///   SENT_NUM_DATABOXES_D: USINT := 5;
///
///END_VAR
///
/// 
///
///PROGRAM OsIniProc
///
///   VAR
///
///		sent_dataBox_as: ARRAY[1..SENT_NUM_DATABOXES_D] OF bds_in_sent_SDDataBox_ts;
///		
///		Init_flag_u8:USINT:=0;	 
///
///   END_VAR
///  
///IF(Init_flag_u8=0) THEN (*To make api call once in application*)
///
///	(* register slow databox *)
///	
///	bds_in_sent_registerSDDataboxes(bds_in_sent_signal_te.K57, ADR(sent_dataBox_as), SENT_NUM_DATABOXES_D);
///	
///	Init_flag_u8:=1;
///  
///END_IF
///
///============================================================================
{attribute 'external_name' := 'cmp_rts_bds_in_sent_registerSDDataboxes'}
FUNCTION bds_in_sent_registerSDDataboxes : USINT
VAR_INPUT
	///The signal name that is assigned to the respective pin configured as SENT input
	signal_e: UINT;
	///Pointer to the message data of type |bds_in_sent_SDDataBox_ts|
	mem_pas: POINTER TO bds_in_sent_SDDataBox_ts;
	/// number of receive databoxes
	num_u8: USINT;
END_VAR

END_FUNCTION

// I/O API/IN legacy/API/bds_in_sent_initSDDatabox
///It initializes a slow serial databox for a particular message of a SENT channel. 
///
///=======
/// Remarks:
///=======
///   + The use of receive databoxes is optional.
///   + Before using this function the receive databoxes must be registered with |bds_in_sent_registerSDDataboxes|  
///   + Each receive databox has to be initialized before it can be used.
///   + By default no databoxes are registered. 
///   + Duplication of same ID should be avoided. 
///
///----------
/// FFI:
///----------
///This API can be used in trusted partitions only. See Freedom from Interference (FFI) concept for more details.
///  
///==================================================================		  			===================================================================================================
///Return value    								  									Description
///==================================================================		  			===================================================================================================
///0																					No error
///1																					Invalid parameter
///2																					New buffer overlaps a present buffer
///3																					A Databox with this id is initialized already
///
///==================================================================		   			===================================================================================================
///
///=======
///Code Example:
///=======
///============================================================================
///
///VAR_GLOBAL CONSTANT
///
///   SENT_NUM_DATABOXES_D: USINT := 5;
///
///   SENT_DATABOX_BUFLEN_D: UDINT := 10;
///
///END_VAR
///
/// 
///
///PROGRAM PLC_PRG OsIniProc
///
///   VAR
///
///		sent_dataBox_as: ARRAY[1..SENT_NUM_DATABOXES_D] OF bds_in_sent_SDDataBox_ts;
///		
///		sent_slowData1_as: ARRAY[1..SENT_DATABOX_BUFLEN_D] OF bds_in_sent_slowData_ts;
///		
///		Init_flag_u8:USINT:=0;	 
///
///   END_VAR
///  
///IF(Init_flag_u8=0) THEN (*To make api call once in application*)
///	
///	(* register slow databox *)
///	
///	bds_in_sent_registerSDDataboxes(bds_in_sent_signal_te.K52, ADR(sent_dataBox_as), SENT_NUM_DATABOXES_D);
///	
///	
///	
///	(* initialize the databox *)
///	
///	bds_in_sent_initSDDatabox(bds_in_sent_signal_te.K52, 1, 2, ADR(sent_slowData1_as), 5);
///	
///	Init_flag_u8:=1;
///  
///END_IF
///
///
///============================================================================
{attribute 'external_name' := 'cmp_rts_bds_in_sent_initSDDatabox'}
FUNCTION bds_in_sent_initSDDatabox : USINT
VAR_INPUT
	///The signal name that is assigned to the respective pin configured as SENT input
	signal_e: UINT;
	///Number of data box
	numDatabox_u8: USINT;
	///Message identifier 
	MsgID_u8: USINT;
	///Pointer to the message data of type |bds_in_sent_slowData_ts|
	buf_pas: POINTER TO bds_in_sent_slowData_ts;
	///length of buffer
	buf_len_u16: UINT;
END_VAR

END_FUNCTION

// I/O API/IN legacy/API/bds_in_sent_getStatus
///Provides the status and error information of a specified SENT channel.
///
///=======
/// Remarks:
///=======
///   + The Error Line Low is set if there is a short circuit to ground (SCG).
///   + The Error Line High is set if there is a open channel or short circuit to battery (SCB).
///   + As soon as the one frame of the FastData (FD) and SlowDat a(SD) is received then the One Frame and One Slow frame received bits will be set.
///   + If the functions |bds_in_sent_getFD| and |bds_in_sent_getSD| are used for reading the FD and SD respectively and a new frame of FD and SD is received then the New Frame and New Slow Frame Received bits will be set. If there is no error then the status information will be 16#3F.
///   + If the FIFO for FD and Databox for SD is registered and a new frame of FD and SD is received, then the New Frame and New Slow Frame Received bits will be set.But since the FIFO and Databox is used these bits will be cleared as soon as the New Frames are received and copied into the FIFO and Databox.So if there is no error then the status information will be 16#17.
///
///
///----------
/// FFI:
///----------
///This API can be used in trusted partitions only. See Freedom from Interference (FFI) concept for more details.
///
///==========================================		  			==========================================		  			================================================
///Value(bit position)   								  		Define														Meaning
///==========================================		  			==========================================		  			================================================
///0															SENT_ERR_NO_ERRORS_DU16										No error
///16#00000001													SENT_STATUS_DRIVER_INIT_DU32								Driver initialized
///16#00000002													SENT_STATUS_DRIVER_RUNNING_DU32            					Driver running
///16#00000004													SENT_STATUS_ONE_FRAME_RECEIVED_DU32 						One frame received
///16#00000008													SENT_STATUS_NEW_FRAME_RECEIVED_DU32 						New frame received
///16#00000010													SENT_STATUS_ONE_SLOW_FRAME_RECEIVED_DU32  					One slow frame received
///16#00000020													SENT_STATUS_NEW_SLOW_FRAME_RECEIVED_DU32   					New slow frame received
///16#00000040													SENT_ERROR_LINE_LOW_DU32                    				Line low   (SCG)
///16#00000080													SENT_ERROR_LINE_HIGH_DU32									Line High (SCB or open channel )
///16#00000100													SENT_ERROR_NODAT_DU32                      					No data received
///16#00000200													SENT_ERROR_NOSIG_DU32										No edges detected
///16#00000400													SENT_ERROR_NOISE_DU32										Noise detected
///16#00000800													SENT_ERROR_DEBOUNCING_DU32  								Debouncing
///16#00001000													SENT_ERROR_CRC_DU32                       					CRC error
///16#00002000													SENT_ERROR_RANGE_DU32                     					Nibble range error
///16#00004000													SENT_ERROR_MISSING_NIBBLE_DU32            					Missing nibble
///16#00008000													SENT_ERROR_TOOMANY_NIBBLES_DU32 							Too many nibbles
///16#00010000													SENT_ERROR_MSG_LOST_DU32                  					Message lost
///16#00020000													SENT_ERROR_SLOW_CRC_DU32                  					Slow channel CRC error
///16#00040000													SENT_ERROR_SLOW_MISSING_FRAME_DU32        					Slow channel missing frame
///16#00080000													SENT_ERROR_NOSLOWDAT_DU32                 					Slow channel no data received
///16#00100000													SENT_ERROR_CAL_PULSE_RANGE_DU32           					Calibration pulse out of range
///16#00200000													SENT_ERROR_CAL_SUCCESSIVE_DEVIATION_DU32  					Calibration pulse successive deviation
///16#00400000													SENT_WARNING_CAL_DEVIATION_20PCT_DU32    					 N/A
///16#00800000													SENT_ERROR_PAUSE_PULSE_RANGE_DU32 							Pause pulse out of range
///16#01000000													SENT_ERROR_FAST_DATA_CTR_DU32 								Fast data counter error
///16#02000000													SENT_ERROR_FAST_DATA_INV_MSN0_DU32							Fast data inverted nibble error
///16#FC000000													RESERVED													N/A
///
///==========================================		  			==========================================					================================================
///
///
/// 
///==================================================================		  			===================================================================================================
///Return value    								  									Description
///==================================================================		  			===================================================================================================
///0																					No error
///1																					Invalid parameter
///2																					Channel is not running
///
///==================================================================		   			===================================================================================================
///
///=======
///Code Example:
///=======
///============================================================================
///
///PROGRAM appl_10ms_task
///
///   VAR
///
///     status_u32: UDINT := 16#00;
///
///   END_VAR
///
///   bds_in_sent_getStatus(bds_in_sent_signal_te.K52,ADR(status_u32));
///
///END
///
///============================================================================
{attribute 'external_name' := 'cmp_rts_bds_in_sent_getStatus'}
FUNCTION bds_in_sent_getStatus : USINT
VAR_INPUT
	///The signal name that is assigned to the respective pin configured as SENT input
	signal_e: UINT;
	///Address where the value is stored.
	value_pu32: POINTER TO UDINT;
END_VAR

END_FUNCTION

// I/O API/IN legacy/API/bds_in_sent_getFD
///Provides the latest received Fast Data of a specified SENT channel.
///
///=======
/// Remarks:
///=======
///   + First check the return value before accessing the message.
///   + Error Handling is done for wrong parameter configuration.
///   + If already fast data FIFO has been registered using the |bds_in_sent_registerFDFifo|,  then the return value FD FIFO register exists. Hence |bds_in_sent_copyFDFifo| should be used to get the FD FIFO.
///   + If the optional decoding fast data is not configured or if the decoding fast data could not happen properly, then the variables in the structure bds_in_sent_decodedFD_ts contain "0".
///   
///
///----------
/// FFI:
///----------
///This API can be used in trusted partitions only. See Freedom from Interference (FFI) concept for more details.
///   
///==================================================================		  			===================================================================================================
///Return value    								  									Description
///==================================================================		  			===================================================================================================
///0																					No error
///1																					Invalid parameter
///2																					Channel is not running
///3																					FD FIFO register exists
///4																					No new FD frame received
///
///==================================================================		   			===================================================================================================
///
///=======
///Code Example:
///=======
///============================================================================
///
///PROGRAM appl_10ms_task
///
///   VAR
///   
///     FD_msg_s: bds_in_sent_decodedFD_ts;
///	 
///     statusFD_u8: USINT := 16#00;
///	 
///   END_VAR
///
///  statusFD_u8 := bds_in_sent_getFD(bds_in_sent_signal_te.K52, ADR(FD_msg_s));
///  
///
///  IF (0 = statusFD_u8) THEN
///  
///    (* Fast Data is valid *)
///	
///  END_IF
///END
///
///============================================================================
{attribute 'external_name' := 'cmp_rts_bds_in_sent_getFD'}
FUNCTION bds_in_sent_getFD : USINT
VAR_INPUT
	///The signal name that is assigned to the respective pin configured as SENT input
	signal_e: UINT;
	///Storage address of the value.
	data_ps: POINTER TO bds_in_sent_decodedFD_ts;
END_VAR

END_FUNCTION

// I/O API/IN legacy/API/bds_in_sent_registerFDFifo
///It registers a fast-data (FD) databox for a SENT channel. The application has to reserve the memory for databox. Further, the databox is managed by the BSW.  
///
///=======
/// Remarks:
///=======
///
///   + The use of receive FD FIFO is optional.
///   + For each SENT channel separate FD FIFO must be registered. 
///   + Only allowed in function OsIniProc().
///   + Please register FIFO only as much as needed. Each FIFO increases the system load. 
///   + Duplication of same buffer register need to be avoided.
/// 
///
///----------
/// FFI:
///----------
///This API can be used in trusted partitions only. See Freedom from Interference (FFI) concept for more details.
///
///==================================================================		  			===================================================================================================
///Return value    								  									Description
///==================================================================		  			===================================================================================================
///0																					No error
///1																					Invalid parameter
///2																					new buffer overlaps a present buffer
///
///==================================================================		   			===================================================================================================
///
///=======
///Code Example:
///=======
///============================================================================
///
///VAR_GLOBAL CONSTANT
///
///   SENT_FD_FIFONUM_D: USINT := 20;
///
///END_VAR
///
/// 
///
///PROGRAM OsIniProc
///
///   VAR
///
///		sent_FDFifo_as: ARRAY[1..SENT_FD_FIFONUM_D] OF bds_in_sent_decodedFD_ts;
///		
///		Init_flag_u8:USINT:=0;	 
///
///   END_VAR
///  
///IF(Init_flag_u8=0) THEN (*To make api call once in application*)
///
///	
///	(* register FastData FIFO *)
///	
///	bds_in_sent_registerFDFifo(bds_in_sent_signal_te.K57, ADR(sent_FDFifo_as[1]), SENT_FD_FIFONUM_D);
///	
///	Init_flag_u8:=1;
///  
///END_IF
///
///
///============================================================================
{attribute 'external_name' := 'cmp_rts_bds_in_sent_registerFDFifo'}
FUNCTION bds_in_sent_registerFDFifo : USINT
VAR_INPUT
	///The signal name that is assigned to the respective pin configured as SENT input
	signal_e: UINT;
	///Pointer to the message data of type |bds_in_sent_decodedFD_ts|
	data_ps: POINTER TO bds_in_sent_decodedFD_ts;
	///size of FIFO
	sizeFifo_u8: USINT;
END_VAR

END_FUNCTION

// I/O API/IN legacy/API/bds_in_sent_copyFDFifo
///This function provides the oldest fast data from a particular FIFO of the specified SENT channel. 
///
///=======
/// Remarks:
///=======
///   + Registration of a FIFO by function |bds_in_sent_registerFDFifo| is essential!
///   + Received fast data of registered FIFO  are saved and can be read by using this function.
///   + First check the return value before accessing the data/message.
///   + Length of copy buffer needs to be greater or equal to the length of the buffer in the |bds_in_sent_registerFDFifo|.
///   
/// 
///----------
/// FFI:
///----------
///This API can be used in trusted partitions only. See Freedom from Interference (FFI) concept for more details.
///  
///==================================================================		  			===================================================================================================
///Return value    								  									Description
///==================================================================		  			===================================================================================================
///0																					No error
///1																					Invalid parameter
///2																					Copy buffer is to small
///3																					Address is invalid
///4																					Buffer is empty
///5																					Buffer overflow error
///6																					Copy data error
///
///==================================================================		   			===================================================================================================
///
///=======
///Code Example:
///=======
///============================================================================
///
///VAR_GLOBAL CONSTANT
///
///   SENT_FD_FIFONUM_D: USINT := 20;
///   
///END_VAR
///
///PROGRAM PLC_PRG
///   VAR
///   
///		sent_FDFifo_as: ARRAY[1..SENT_FD_FIFONUM_D] OF bds_in_sent_decodedFD_ts;
///		
///		sent_FDfifoCopy: ARRAY[1..SENT_FD_FIFONUM_D] OF bds_in_sent_decodedFD_ts;
///		
///		sent_copy: bds_in_sent_copyFDBuf_ts;
///		
///		Init_flag_u8:USINT:=0;
///	 
///   END_VAR
///   
///IF(Init_flag_u8=0) THEN (*To make api call once in application*)
///		
///	(* register fast Data fifo *)
///	
///	bds_in_sent_registerFDFifo(bds_in_sent_signal_te.K52, ADR(sent_FDFifo_as[1]), SENT_FD_FIFONUM_D);
///	
///	(* copy register fast Data fifo *)
///	
///	bds_in_sent_registerCopyFDFifo(ADR(sent_copy), ADR(sent_FDfifoCopy), SENT_FD_FIFONUM_D);
///	
///	sent_copy.start_pas := sent_FDfifoCopy;
///	
///	sent_copy.lengthCopyBuf_u8 := 20;
///	
///	Init_flag_u8:=1;
///  
///END_IF
///
///PROGRAM appl_10ms_task
///VAR
///
///  statusFDFIFO_u8 : USINT;
///  statusFDFIFO_u8 := bds_in_sent_copyFDFifo(bds_in_sent_signal_te.K52, ADR(sent_copy));
///
/// 
///END_VAR
///
///
///IF (0 = statusFDFIFO_u8) THEN
///
///	(* Message in structure sent_copy is valid *)
///	
///END_IF
///
///
///============================================================================
{attribute 'external_name' := 'cmp_rts_bds_in_sent_copyFDFifo'}
FUNCTION bds_in_sent_copyFDFifo : USINT
VAR_INPUT
	///The signal name that is assigned to the respective pin configured as SENT input
	signal_e: UINT;
	///pointer to |bds_in_sent_copyFDBuf_ts|
	data_ps: POINTER TO bds_in_sent_copyFDBuf_ts;
END_VAR

END_FUNCTION

// I/O API/IN legacy/API/bds_in_sent_registerCopyFDFifo
///The function registers the copy buffer for fast data FIFO for specified SENT channel. 
///
///=======
/// Remarks:
///=======
///
///   + A copy buffer must be registered with a number of FD Fifo data. The number must be equal with the maximum number of FD FIFO data which are registered for the buffers using |bds_in_sent_registerFDFifo|.
///   + Please register the copy buffer for fast data FIFO only as much as needed, because each registered copy buffer for fast data FIFO increases the system load.
///   + The application must define the buffer info structure and the buffer (memory space).
///   + For access to the FD FIFO data the function |bds_in_sent_copyFDFifo| is used.
/// 
///----------
/// FFI:
///----------
///This API can be used in trusted partitions only. See Freedom from Interference (FFI) concept for more details.
/// 
///==================================================================		  			===================================================================================================
///Return value    								  									Description
///==================================================================		  			===================================================================================================
///0																					No error
///1																					Invalid parameter
///2																					new buffer overlaps a present buffer
///
///==================================================================		   			===================================================================================================
///
///=======
///Code Example:
///=======
///============================================================================
///
///VAR_GLOBAL CONSTANT
///
///   SENT_FD_FIFONUM_D: USINT := 20;
///
///END_VAR
///
/// 
///
///PROGRAM PLC_PRG
///
///   VAR
///
///		sent_FDFifo_as: ARRAY[1..SENT_FD_FIFONUM_D] OF bds_in_sent_decodedFD_ts;
///		
///		sent_FDfifoCopy: ARRAY[1..SENT_FD_FIFONUM_D] OF bds_in_sent_decodedFD_ts;
///		
///		sent_copy: bds_in_sent_copyFDBuf_ts;
///		
///		Init_flag_u8:USINT:=0;	 
///
///   END_VAR
///  
///IF(Init_flag_u8=0) THEN (*To make api call once in application*)
///
///	(* register fast Data fifo *)
///	
///	bds_in_sent_registerFDFifo(bds_in_sent_signal_te.K52, ADR(sent_FDFifo_as[1]), SENT_FD_FIFONUM_D);
///	
///	(* copy register fast Data fifo *)
///	
///	bds_in_sent_registerCopyFDFifo(ADR(sent_copy), ADR(sent_FDfifoCopy), SENT_FD_FIFONUM_D);
///	
///	Init_flag_u8:=1;
///  
///END_IF
///
///============================================================================
{attribute 'external_name' := 'cmp_rts_bds_in_sent_registerCopyFDFifo'}
FUNCTION bds_in_sent_registerCopyFDFifo : USINT
VAR_INPUT
	///pointer to |bds_in_sent_copyFDBuf_ts|
	sent_copyFDBufInfo_ps: POINTER TO bds_in_sent_copyFDBuf_ts;
	///pointer to |bds_in_sent_decodedFD_ts|
	buf_ps: POINTER TO bds_in_sent_decodedFD_ts;
	///length of FIFO.
	lenFifo_u8: USINT;
END_VAR

END_FUNCTION

// I/O API/IN legacy/API/bds_in_sent_getSD
///Provides the latest received Slow Data of a specified SENT channel.
///
///=======
/// Remarks:
///=======
///   + First check the return value before accessing the message.
///   + Error Handling is done for wrong parameter configuration.
///   + If slow databox has already been configured using the |bds_in_sent_registerSDDataboxes|, then the return value SD Databox register exists. Hence |bds_in_sent_getSDDatabox|  should be used to get the SD Databox.
///
///----------
/// FFI:
///----------
///This API can be used in trusted partitions only. See Freedom from Interference (FFI) concept for more details.
///   
///==================================================================		  			===================================================================================================
///Return value    								  									Description
///==================================================================		  			===================================================================================================
///0																					No error
///1																					Invalid parameter
///2																					SENT channel is not running
///3																					SD Databox register exists
///4																					No new SD frame received
///
///==================================================================		   			===================================================================================================
///
///=======
///Code Example:
///=======
///============================================================================
///
///PROGRAM appl_10ms_task
///
///   VAR
///   
///     SD_msg_s: bds_in_sent_slowData_ts;
///	 
///     statusSD_u8: USINT := 16#00;
///	 
///   END_VAR
///
///  statusSD_u8 := bds_in_sent_getSD(bds_in_sent_signal_te.K52, ADR(SD_msg_s));
///
///  IF (0 = statusSD_u8) THEN
///  
///    (* slow data is valid *)
///	
///  END_IF
///
///============================================================================
{attribute 'external_name' := 'cmp_rts_bds_in_sent_getSD'}
FUNCTION bds_in_sent_getSD : USINT
VAR_INPUT
	///The signal name that is assigned to the respective pin configured as SENT input
	signal_e: UINT;
	///Storage address of the value.
	data_ps: POINTER TO bds_in_sent_slowData_ts;
END_VAR

END_FUNCTION

// System API/DSM/API/Macro Functions/bds_dsm_DFC_da
///It returns the debounce activ bit fields from DFC status word
{attribute 'external_name' := 'cmp_rts_bds_dsm_DFC_da'}
FUNCTION bds_dsm_DFC_da : USINT
VAR_INPUT
	dfc_u16: UINT;
END_VAR

END_FUNCTION

// I/O API/OUT_LEGACY/bds_out_po_cfgPeriod
///Reconfigures the period [µs] of the proportional output.
///
///=======
/// Remarks:
///=======
///
///   + For the low power outputs the period range is from from 300 to 31000µs.
///   + For the high power outputs the period range is from 1000us to 100000µs and for low side  4000 to 100000µs and only multiples of 1000µs are accepted.
///   + For more information see |bds_out_po_getStatus|.
///   + The structure member status_b16 holds the information regarding the configuration.
///   + This function should be called only once in the application.
///
///----------
/// FFI:
///----------
///This API can be used in trusted partitions  For untrusted partitions use |bds_out_po_cfgPeriod_ffi|. See Freedom from Interference (FFI) concept for more details.
///
///==================================================================		  			===================================================================================================
///Return value    								  									Description
///==================================================================		  			===================================================================================================
///0																					No error.
///1																					A parameter is invalid.
///2																					Function call was erroneous.
///
///==================================================================		   			===================================================================================================
///
///=======
///Code Example:
///=======
///============================================================================
///
///PROGRAM PLC_PRG
///
///VAR
///
///	Init_flag_u8:USINT:=0;
///
///END_VAR
///  
///IF(Init_flag_u8=0) THEN (*To make api call once in application*)
///				
///	(* configure a period of 20ms for output K73 *)
///	
///	bds_out_po_cfgPeriod(bds_out_po_signal_te.K73, 20000);
///  
///	Init_flag_u8:=1;
///  
///END_IF
///
///============================================================================
{attribute 'external_name' := 'cmp_rts_bds_out_po_cfgPeriod'}
FUNCTION bds_out_po_cfgPeriod : USINT
VAR_INPUT
	///The connector assigned signal name of the output.
	signal_e: UINT;
	///New period [µs].Range:
	///   + Low power output: 300 to 31000
	///   + High power output high side: 1000, 4000, 5000 to 100000
	///   + High power output low side: 4000, 5000 tp 100000
	///
	///Note:For the high power outputs are only multiples of 1ms allowed.
	period_u32: UDINT;
END_VAR

END_FUNCTION

// I/O API/OUT/FFI_API/bds_out_po_cfgPeriod_ffi
{attribute 'external_name' := 'cmp_rts_bds_out_po_cfgPeriod_ffi'}
FUNCTION bds_out_po_cfgPeriod_ffi : USINT
VAR_INPUT
	///The connector assigned signal name of the output.
	signal_e: UINT;
	///New period [µs].Range:
	///   + Low power output: 300 to 31000
	///   + High power output high side: 1000, 4000, 5000 to 100000
	///   + High power output low side: 4000, 5000 tp 100000
	///
	///Note:For the high power outputs are only multiples of 1ms allowed.
	period_u32: UDINT;
END_VAR

END_FUNCTION

// I/O API/OUT_LEGACY/bds_out_po_disable
///Disables unused proportional output to avoid faults on unused outputs.
///
///=======
/// Remarks:
///=======
///   + Prevents the setting of open load faults at an unused output..
///   + The output should be disabled during start up.
///   + This function should be called only once in the application.
///
///----------
/// FFI:
///----------
///This API can be used in trusted partitions . For untrusted partitions use |bds_out_po_disable_ffi|. See Freedom from Interference (FFI) concept for more details.
///   
///------
/// Attention:
///------
///
///If an output is  disabled, faults are not longer detected and also the control of the output is suppressed
///
///==================================================================		  			===================================================================================================
///Return value    								  									Description
///==================================================================		  			===================================================================================================
///0																					No error.
///1																					A parameter is invalid.
///2																					Output is already configured as safout, output can't be disabled
///
///==================================================================		   			===================================================================================================
///
///=======
///Code Example:
///=======
///============================================================================
///
///PROGRAM PLC_PRG
///
///VAR
///
///	Init_flag_u8:USINT:=0;
///
///END_VAR
///  
///IF(Init_flag_u8=0) THEN (*To make api call once in application*)
///				
///	(* disable output K83 *)
///	
///	bds_out_po_disable(bds_out_po_signal_te.K83, STD_ON);
///  
///	Init_flag_u8:=1;
///  
///END_IF
///
///============================================================================
{attribute 'external_name' := 'cmp_rts_bds_out_po_disable'}
FUNCTION bds_out_po_disable : USINT
VAR_INPUT
	///The connector assigned signal name of the output.
	signal_e: UINT;
	///The possible states are
	///   + STD_OFF - Enable the output (default)
	///   + STD_ON   - Disable the output
	state_u8: USINT;
END_VAR

END_FUNCTION

// I/O API/OUT/FFI_API/bds_out_po_disable_ffi
{attribute 'external_name' := 'cmp_rts_bds_out_po_disable_ffi'}
FUNCTION bds_out_po_disable_ffi : USINT
VAR_INPUT
	///The connector assigned signal name of the output.
	signal_e: UINT;
	///The possible states are
	///   + STD_OFF - Enable the output (default)
	///   + STD_ON   - Disable the output
	state_u8: USINT;
END_VAR

END_FUNCTION

// Diagnostics API/UDS/API/bds_uds_updNodeIDinNVM
///This function updates Node ID in NVM shared configuration.
///
///=======
/// Remarks:
///=======
///    + This will change the node ID in NVM section, not in the UDS stack.
///    + To read the configured node ID |bds_uds_getNodeID| can be used.
///    + The set node ID will be configured in the UDS stack after one of the following actions,
///	    + |bds_sys_resetECU| is invoked.
///	    + |bds_sys_startLoader| is invoked.
///	    + T15 is switched OFF.
///    + The |GVL_uds| is given for usage of defines.
///
///----------
/// FFI:
///----------
///This API can be used in trusted partitions only. See Freedom from Interference (FFI) concept for more details.
///		
///==================================================================		  			===================================================================================================
///Return value    								  									Description
///==================================================================		  			===================================================================================================
///16#00																				No error
///16#03																				Invalid Node ID
///
///==================================================================		   			===================================================================================================
{attribute 'external_name' := 'cmp_rts_bds_uds_updNodeIDinNVM'}
FUNCTION bds_uds_updNodeIDinNVM : USINT
VAR_INPUT
	///Node ID of UDS stack which has to be configured in the next initialization.
	///    + The possible values are:16#00 to 16#FE
	///    + Default value are :16#01
	nodeId_u8: USINT;
END_VAR

END_FUNCTION

// Diagnostics API/XCP/API/bds_xcp_setMode
///This function sets the mode (Enable/Disable) of XCP.
///
///=======
/// Remarks:
///=======
///
///    + The |GVL_xcp| is given for usage of defines.
///
///----------
/// FFI:
///----------
///This API can be used in trusted partitions only. See Freedom from Interference (FFI) concept for more details.
///
///----------
/// DANGER:
///----------
///
///Software running on the ECU can be manipulated with XCP. That will lead to both a security and a safety risk. Life and health can be endangered. Thus, it must be impossible to use XCP on serial machines.
///
///
///==================================================================		  			===================================================================================================
///Return value    								  									Description
///==================================================================		  			===================================================================================================
///None																				None
///
///==================================================================		   			===================================================================================================
///
///
///=======
///Code Example:
///=======
///============================================================================
///
///PROGRAM PLC_PRG
///  VAR
///  
///  END_VAR
///
///  (* Enable XCP *)
///  
///  bds_xcp_setMode(BDS_ENABLE_XCP_DU16);
///
///============================================================================
{attribute 'external_name' := 'cmp_rts_bds_xcp_setMode'}
FUNCTION bds_xcp_setMode : BOOL
VAR_INPUT
	///Indicates whether XCP should be enabled or disabled.
	///
	///Possible values:
	///    + BDS_DISABLE_XCP_DU16 (16#0000)           : Disable XCP communication.
	///    + BDS_ENABLE_XCP_DU16  (16#FFFF)           : Enable read, write Access in XCP.
	///    + BDS_ENABLE_XCP_READ_DU16 (16#FFFE)           : Enable read only Access in XCP.
	mode_u16: UINT;
END_VAR

END_FUNCTION

// I/O API/IN legacy/API/bds_in_ri
///Provides the resistance of the input.
///
///=======
/// Remarks:
///=======
///   + The used measurement range is defined between 20 ohm to 400k ohm, Also see  |bds_in_ri_cfg| for the configuration of  thresholds for diagnostics.
///   + The possible measurement range is higher than 700k ohm (These are the value for an open load or a short circuit to battery). 
///   + For more information regarding the signal acquisition see Analog voltage acquisition.
///
///
///----------
/// FFI:
///----------
///This API can be used in trusted partitions only. See Freedom from Interference (FFI) concept for more details.
///
///==================================================================		  			===================================================================================================
///Return value    								  									Description
///==================================================================		  			===================================================================================================
///0																					No error
///1																					Invalid parameter
///2																					Function call was erroneous
///
///==================================================================		   			===================================================================================================
///
///=======
///Code Example:
///=======
///============================================================================
///
///PROGRAM appl_10ms_task
///
///  VAR
///  
///    ohmK60_u32: UDINT := 16#00;
///	
///  END_VAR
///
///(* get the resistance of input K60 *)
///
///bds_in_ri(bds_in_ri_signal_te.K60, ADR(ohmK60_u32));
///
///END
///
///============================================================================
{attribute 'external_name' := 'cmp_rts_bds_in_ri'}
FUNCTION bds_in_ri : USINT
VAR_INPUT
	///The signal name that is assigned to the respective pin configured as resistance input
	signal_e: UINT;
	///Storage address of the value.
	///
	///Range:
	///20..400000 [ohm]
	///
	///Value for an open load or a short circuit to battery:
	///> 700000 [ohm]
	value_pu32: POINTER TO UDINT;
END_VAR

END_FUNCTION

// System API/DSM/API/Macro Functions/bds_dsm_DFC_dfl
///It returns the debounced fault level bit fields from DFC status word
{attribute 'external_name' := 'cmp_rts_bds_dsm_DFC_dfl'}
FUNCTION bds_dsm_DFC_dfl : USINT
VAR_INPUT
	dfc_u16: UINT;
END_VAR

END_FUNCTION

// System API/DSM/API/bds_dsm_getErrors
///This function is used to get all DFCs with the specified status.
///
///=======
/// Remarks:
///=======
///    + The |GVL_dsm| is given for usage of defines.
///	
///----------
/// FFI:
///----------
///This API can be used in trusted partitions . For untrusted partitions use |bds_dsm_getErrors_ffi|. See Freedom from Interference (FFI) concept for more details.
///
///==================================================================		  			===================================================================================================
///Return value    								  									Description
///==================================================================		  			===================================================================================================
///16#0000: BDS_DSM_NO_ERROR_DU16														Update Number of Error is successful.
///16#0004: BDS_DSM_INVALID_PTR_DU16													Invalid Pointer
///16#0005: BDS_DSM_MASK_ERROR_DU16													Invalid Mask.
///16#0007: BDS_DSM_INVALID_MAX_ERROR_DU16 											Invalid Max Error.
///16#0008:BDS_DSM_OVERFLOW_ERROR_DU16													Number of error are more than Max Error. 
///16#000C: BDS_DSM_FFI_ACCESS_ERROR_DU16												Invalid Access to FFI variant API call.
///
///==================================================================		   			===================================================================================================
///
///
///=======
///Code Example:
///=======
///============================================================================
///
///PROGRAM DSM
///
///VAR
///
///	mask_s : UINT := BDS_DSM_SET_ACTIVE_ERROR_MASK_DU16;
///
///	startFromBegin_l: BOOL := TRUE;
///
///	maxNum_u16:UINT := 32;
///
///	error_count_u16: UINT;
///
///	dfc_active_as: ARRAY [1..32] OF bds_dsm_dfc_ts;
///
///	status_u16: UINT;
///
///END_VAR
///
///
///(*Get errors*)
///
///status_u16 := bds_dsm_getErrors(mask_s,startFromBegin_l,maxNum_u16,ADR(error_count_u16),ADR(dfc_active_as)); 
///
///IF status_u16 = BDS_DSM_NO_ERROR_DU16 THEN
///
///	(*Number of Errors has been read successfully*)
///
///END_IF
///
///
///============================================================================
///
{attribute 'external_name' := 'cmp_rts_bds_dsm_getErrors'}
FUNCTION bds_dsm_getErrors : UINT
VAR_INPUT
	///The kind of error status can be specified in detail by means of this mask.
	///
	///Possible values:
	///    + BDS_DSM_SET_ACTIVE_ERROR_MASK_DU16 ( 16#18 ) - Fault is active.
	///    + BDS_DSM_SET_TESTED_ONCE_MASK_DU16 ( 16#08 ) - DFC was tested at least once since start or reset.
	///    + BDS_DSM_SET_TESTED_OK_MASK_DU16 ( 16#20 ) - DFC was at least once ok tested since start or reset.  
	///    + BDS_DSM_SET_FAILED_SINCE_CLEAR_MASK_DU16 ( 16#80 ) - Fault occured at least once since error was deleted from memory.
	mask_s: UINT;
	///
	///    + TRUE: Query is started from the beginning of DFES.
	///    + FALSE: Query is continued with the next index where the last query was finished.
	startFromBegin_l: BOOL;
	///Maximal number of errors/DFCs which can be returned.
	maxNum_u16: UINT;
	///Pointer to a variable where the number of errors/DFCs is returned.
	num_pu16: POINTER TO UINT;
	///Pointer to a variable/an array where the errors/DFCs will be returned (note: this array must have the size for the number of errors/DFCs specified in parameter maxNum_u16).
	dfc_ps: POINTER TO bds_dsm_dfc_ts;
END_VAR

END_FUNCTION

// System API/DSM/FFI_API/bds_dsm_getErrors_ffi
{attribute 'external_name' := 'cmp_rts_bds_dsm_getErrors_ffi'}
FUNCTION bds_dsm_getErrors_ffi : UINT
VAR_INPUT
	///The kind of error status can be specified in detail by means of this mask.
	///
	///Possible values:
	///    + BDS_DSM_SET_ACTIVE_ERROR_MASK_DU16 ( 16#18 ) - Fault is active.
	///    + BDS_DSM_SET_TESTED_ONCE_MASK_DU16 ( 16#08 ) - DFC was tested at least once since start or reset.
	///    + BDS_DSM_SET_TESTED_OK_MASK_DU16 ( 16#20 ) - DFC was at least once ok tested since start or reset.  
	///    + BDS_DSM_SET_FAILED_SINCE_CLEAR_MASK_DU16 ( 16#80 ) - Fault occured at least once since error was deleted from memory.
	mask_s: UINT;
	///
	///    + TRUE: Query is started from the beginning of DFES.
	///    + FALSE: Query is continued with the next index where the last query was finished.
	startFromBegin_l: BOOL;
	///Maximal number of errors/DFCs which can be returned.
	maxNum_u16: UINT;
	///Pointer to a variable where the number of errors/DFCs is returned.
	num_pu16: POINTER TO UINT;
	///Pointer to a variable/an array where the errors/DFCs will be returned (note: this array must have the size for the number of errors/DFCs specified in parameter maxNum_u16).
	dfc_ps: POINTER TO bds_dsm_dfc_ts;
END_VAR

END_FUNCTION

// System API/DSM/API/bds_dsm_getDTC_Status
///This function is used to get the 16 bit DTC status word of specified DFC.
///
///=======
/// Remarks:
///=======
///    + The |GVL_dsm| is given for usage of defines.
///    + For information on 16 bit DTC status word refer Diagnostic Fault Check. 
///
///----------
/// FFI:
///----------
///This API can be used in trusted partitions only. See Freedom from Interference (FFI) concept for more details.
///	
///==================================================================		  			===================================================================================================
///Return value    								  									Description
///==================================================================		  			===================================================================================================
///16#0000: BDS_DSM_NO_ERROR_DU16														Update of Status is Successful .
///16#0004: BDS_DSM_INVALID_PTR_DU16													Invalid Pointer.
///16#000B: BDS_DSM_NO_DTC_AVAILABLE_DU16  											Invalid DTC input.
///
///==================================================================		   			===================================================================================================
///
///
///=======
///Code Example:
///=======
///============================================================================
///
///PROGRAM DSM
///
///VAR
///
///	status_u16: UINT;
///
///	dfc_s: bds_dsm_dfc_ts;	
///
///	dfc_ts : DFC_bds_NoDebFault1;
///
///	error_u16:UINT;
///
///END_VAR
///
///dfc_s.id := dfc_ts.DFCid;
///
///(*Deletes the Error status from DFC and related DFES entry*)
///
///error_u16 := bds_dsm_getDTC_Status(dtc_u16, ADR(status_u16));
///
///if error_u16 = BDS_DSM_NO_ERROR_DU16 THEN
///
///	(*Error Status has been reported succesfully*)
///
///END_IF
///
///============================================================================
///
{attribute 'external_name' := 'cmp_rts_bds_dsm_getDTC_Status'}
FUNCTION bds_dsm_getDTC_Status : UINT
VAR_INPUT
	///DTC value : It is configured using easyConfig tool.
	dtc_u16: UINT;
	///Pointer to variable where the 16 bit DTC status word is returned.
	dtc_status: POINTER TO UINT;
END_VAR

END_FUNCTION

